// TwinCAT 3 PLC project TC3_CNCPLCBase
// Title: CNC PLC Project
// Company: Beckhoff Automation GmbH
// Author: Beckhoff Automation GmbH
// ProjectVersion: 3.1.5000.18
// Description: TwinCAT CNC Base Project
// ProgramVersion: 3.1.4026.23
// libraries:
//   Tc2_CncHli, * (Beckhoff Automation GmbH)
//   Tc2_Standard, * (Beckhoff Automation GmbH)
//   Tc2_System, * (Beckhoff Automation GmbH)
//   Tc3_CNC, * (Beckhoff Automation GmbH)
//   Tc3_EventLogger, * (Beckhoff Automation GmbH)
//   Tc3_JsonXml, * (Beckhoff Automation GmbH)
//   Tc3_Module, * (Beckhoff Automation GmbH)
// project tree:
//   CNC/ Global_CNC.TcGVL, PRG_CNCAxesHandler.TcPOU, PRG_CNCChannelHandler.TcPOU, PRG_CNCDiagnostics.TcPOU, PRG_CNCManualMode.TcPOU, PRG_CNCVariablesViewer.TcPOU, PRG_ManualFnc.TcPOU
//   / FAST.TcPOU, MAIN.TcPOU, PlcFastTask.TcTTO, PlcTask.TcTTO
//   HMI/ Global_HMI.TcGVL, ST_MachineData.TcDUT, ST_MachineMode.TcDUT, ST_MANUAL.TcDUT, ST_Position.TcDUT
//   Messages/ FB_Alarm.TcPOU, Global_Messages.TcGVL, PRG_MessagesV2.TcPOU
//   Samples/ PRG_FastMFunctions.TcPOU
// real-time tasks:
//   TASK PlcTask: cycle T#10ms, priority 20, ADS port 350
//   TASK PlcFastTask: cycle T#10ms, priority 21, ADS port 351
//   TASK CNC-Task ADS: cycle default, priority 7, ADS port 558
//   TASK CNC-Task COM: cycle T#10ms, priority 13, ADS port 556
//   TASK CNC-Task SDA: cycle T#10ms, priority 8, ADS port 555
//   TASK CNC-Task GEO: cycle T#2ms, priority 3, ADS port 554

CONFIGURATION TC3_CNCPLCBase
    RESOURCE PLC ON TwinCAT3
        TASK PlcFastTask(INTERVAL := T#10ms, PRIORITY := 21);
        TASK PlcTask(INTERVAL := T#10ms, PRIORITY := 20);
        PROGRAM FAST WITH PlcFastTask : FAST;
        PROGRAM MAIN WITH PlcTask : MAIN;
    END_RESOURCE
END_CONFIGURATION

// ---- HMI/ST_MachineData.TcDUT
TYPE ST_MachineData :
STRUCT
	// @1: Value1
	Value1: INT;
	// @1: Bool Value
	Value2: bool;
	// @1: Position
	pos : ST_Position;
	// @1: Manual @6:1
	manualFunction : ST_Manual;
END_STRUCT
END_TYPE

// ---- HMI/ST_MachineMode.TcDUT
TYPE ST_MachineMode :
STRUCT
	/// Operation Mode 
	Standby: BOOL;
	Manual: BOOL;
	MDI: BOOL;
	Automatic: BOOL;
	///REFERENCE		: BOOL;  TC3HR
	Homing: BOOL;
	/// Operation State
	Select : BOOL; 
	Ready  : BOOL;
	Start: BOOL;
	Stop: BOOL;
	Reset: BOOL;
	Error: BOOL;
	/// Special functions 
	ChannelSignals: ST_ChannelSignals;
	BlockSearch: ST_BlockSearch;
	SyntaxCheck: ST_SyntaxCheck;
	ManualMode: ST_ManualMode;
	/// Strings 
//	ProgramName: STRING(1024);
//	MDIString: STRING(1024);
	ProgramName: STRING(HLI_IMCM_MODE_STATE_PARAM_STRL);
	MDIString: STRING(HLI_IMCM_MODE_STATE_PARAM_STRL);

END_STRUCT
END_TYPE

// ---- HMI/ST_MANUAL.TcDUT
TYPE ST_MANUAL :
STRUCT
	// @1:cylinder one @2:on:1 @3:off:1 @4:pos1:1 @5:pos2:0
	cyl1 			: BYTE;	
	cyl1Status		: BYTE;
	
	// @1:conveyor @2:IMG1:1 @2:IMG2 @3:IMG15 @4:IMG16 @5:IMG7 @6:IMG13 @7:IMG14
	conv 			: BYTE;
	convStatus 		: BYTE;
	
	
END_STRUCT
END_TYPE

// ---- HMI/ST_Position.TcDUT
TYPE ST_Position :
STRUCT
	// @1:X
	x	:	LREAL;
	// @1:Y
	y	: 	LREAL;
	// @1:Z	
	Z	: 	LREAL;
END_STRUCT
END_TYPE

// ---- CNC/Global_CNC.TcGVL
VAR_GLOBAL CONSTANT
	MAX_USED_CHANNEL_IDX		: INT := 2;									(* Max index of channel that is used starting at 0, example: 1 -> totally 2 channels, maximum of 11 (12 channels) is allowed here *)
	libVersion					: ST_LibVersion := stLibVersion_Tc3_CNC;  	 
END_VAR

// ---- HMI/Global_HMI.TcGVL
VAR_GLOBAL
	/// HMI -> PLC 
	PLCChannelSignals: ST_ChannelSignals;
	/// HMI -> PLC 
	PLCSelectedChannel: INT := 0;
	/// HMI -> PLC 
	PLCFeedOverride: UINT := 100;
	/// HMI -> PLC 
	PLCSpindleOverride: UINT := 100;
	/// HMI -> PLC 
	PLCAxisEnable: BOOL;
	/// PLC -> HMI  
	PLCStatusAxisEnabled : BOOL;	
	/// HMI -> PLC 
	PLCReset: BOOL;
	PLCMachineMode: ARRAY[0..MAX_USED_CHANNEL_IDX] OF ST_MachineMode;
	/// PLC -> HMI : angewähltes File 
	PLCToHmiFile: STRING(255);
	/// Variablen für das Module "InformPlc" 
	bToggle: BOOL;
	sActualForm: STRING(255);
	nUserLevel: INT;
	sUserName: STRING(255);
	/// steigende Flanke: Applikation beenden 
	bExitApp: BOOL;	
	
	userActivity : BOOL;
	
	// @1:MachineData
	MachineData : ST_MachineData;
	
	// spindle manual mode
	nSpindleRpm:	DINT;	
	bSpindleStart: BOOL;
	bSpindleStop: BOOL;
	
	ManualFnc : ARRAY[0..3] OF FB_ManualFncFull;
	
END_VAR

// ---- Messages/Global_Messages.TcGVL
VAR_GLOBAL
	///--------------------------
	///	Messages                
	///--------------------------
	MSG_WARNING_List: ARRAY[FIRST_MESSAGE..LAST_MESSAGE] OF BOOL;
	MSG_WARNING_ListQuit: ARRAY[FIRST_MESSAGE..LAST_MESSAGE] OF BOOL;	
	MSG_ALARM_List: ARRAY[FIRST_MESSAGE..LAST_MESSAGE] OF BOOL;
	MSG_ALARM_ListQuit: ARRAY[FIRST_MESSAGE..LAST_MESSAGE] OF BOOL;			
END_VAR

VAR_GLOBAL CONSTANT
	FIRST_MESSAGE: UDINT := 1;
	LAST_MESSAGE: UDINT := 50;	
END_VAR

// ---- FAST.TcPOU
PROGRAM FAST
VAR
	nChan : INT;
	MOS_TS: INT;
	i: INT;	
	ChannelMHTFunction : ARRAY[0..MAX_USED_CHANNEL_IDX] OF HLI3_QuitChannelMHTFunction;
END_VAR

(****************************************************************************************)
(*	  							Wait for HLI initialization								*)
(****************************************************************************************)
IF NOT CNCSystem.bHLIInit THEN
	RETURN;
END_IF

IF PRG_CNCChannelHandler.stOptions.bDisableMFunctHandling THEN
	FOR i := 0 TO MAX_USED_CHANNEL_IDX DO
		ChannelMHTFunction[i](nChanIdx:=0, bM30Acknowledgement := TRUE);
	END_FOR
END_IF	

(* Programm call for MOS_TS M functions *)
// PRG_FastMFunctions();

END_PROGRAM

// ---- CNC/PRG_CNCChannelHandler.TcPOU
PROGRAM PRG_CNCChannelHandler
VAR	
	nChan					: INT;
	nOldSelectedChannel		: UDINT;
	CNCChannel				: ARRAY[0..MAX_USED_CHANNEL_IDX] OF HLI3_CNCChannel;	
	BlockSearch_Channel		: ARRAY[0..MAX_USED_CHANNEL_IDX] OF HLI3_BlockSearch;
	ErrorHandler_Channel	: ARRAY[0..MAX_USED_CHANNEL_IDX] OF FB_ChannelError;
	nChanNo: UDINT;	
	i: INT;	
	stOptions				: ST_CNC_CH_Options;
END_VAR

(****************************************************************************************)
(* POU:		PRG_ChannelHandler                     										*)
(* Type:	PRG																			*)
(* Author: 	HR / TV / MiB                                          						*)
(* Date: 	23.01.11																	*)
(* Last:	29.03.18																	*)
(* Rev.: 	1.6                                              							*)
(* ------------------------------------------------------------------------------------ *)
(* Desc:	Description																	*)
(****************************************************************************************)

(****************************************************************************************)
(*	  Map CNC function selection from HMI to selected channel (and state vice versa)  	*)
(****************************************************************************************)
IF (nOldSelectedChannel <>INT_TO_UDINT(PLCSelectedChannel)) THEN
	PLCChannelSignals.SingleBlock 		:= PLCMachineMode[PLCSelectedChannel].ChannelSignals.SingleBlock;
	PLCChannelSignals.PrgBlockIgnore	:= PLCMachineMode[PLCSelectedChannel].ChannelSignals.PrgBlockIgnore;
	PLCChannelSignals.M01Stop 			:= PLCMachineMode[PLCSelectedChannel].ChannelSignals.M01Stop;
	PLCChannelSignals.Backward 			:= PLCMachineMode[PLCSelectedChannel].ChannelSignals.Backward;
	PLCChannelSignals.FeedHold 			:= PLCMachineMode[PLCSelectedChannel].ChannelSignals.FeedHold;
	nOldSelectedChannel 				:= INT_TO_UDINT(PLCSelectedChannel);
END_IF

PLCMachineMode[PLCSelectedChannel].ChannelSignals.SingleBlock 		:= PLCChannelSignals.SingleBlock;
PLCMachineMode[PLCSelectedChannel].ChannelSignals.PrgBlockIgnore 	:= PLCChannelSignals.PrgBlockIgnore;
PLCMachineMode[PLCSelectedChannel].ChannelSignals.M01Stop 			:= PLCChannelSignals.M01Stop;
PLCMachineMode[PLCSelectedChannel].ChannelSignals.Backward 		:= PLCChannelSignals.Backward;
PLCMachineMode[PLCSelectedChannel].ChannelSignals.FeedHold 		:= PLCChannelSignals.FeedHold;


stOptions.bReferenceModeStartRequired := FALSE;

FOR i := 0 TO MAX_USED_CHANNEL_IDX DO
		
	nChan := i;	
	IF (HLI3_CheckChannelValid(nChan)) THEN		
		
		(* Error handler for channel 1 *)
		ErrorHandler_Channel[nChan](nChanIdx			:= nCHan);				
				
		(* Channel interface *)
		CNCChannel[nChan]
			(nChanIdx			:= nChan,							
			 // Operation Mode with VAR_IN_OUT Variables 
			 bModeStandby		:= PLCMachineMode[nChan].Standby,
			 bModeAutomatic		:= PLCMachineMode[nChan].Automatic,
			 bModeManual		:= PLCMachineMode[nChan].Manual,
			 bModeMDI			:= PLCMachineMode[nChan].MDI,	 
			 bModeReference		:= PLCMachineMode[nChan].Homing,
			 // Operation State with VAR_IN_OUT Variables
			 bStateSelect		:= PLCMachineMode[nChan].Select,
			 bStateReady		:= PLCMachineMode[nChan].Ready,
			 bStateStart		:= PLCMachineMode[nChan].Start,
			 bStateStop			:= PLCMachineMode[nChan].Stop,
			 bStateReset		:= PLCMachineMode[nChan].Reset,
			 // Operation Mode with VAR_IN Varaibles, the command is executed with a rising edge 
			 bCmdAutomatic 		:= FALSE,
			 bCmdManual 		:= FALSE,
    		 bCmdReference 		:= FALSE,
    		 bCmdMDI 			:= FALSE,		
			 // Operation State with VAR_IN Varaibles, the command is executed with a rising edge
			 bCmdStart 			:= FALSE,
			 bCmdStop  			:= FALSE,
	         bCmdReset 			:= FALSE,					 			 
			 // EmergencyStop 
			 bEmergencyStop 	:= FALSE,		(* If TRUE the interpolation will be aborted, Signal is no TwinSAFE function !*)
			 // Override 
			 nFeedOverride		:= PLCFeedOverride * 10,
			 nRapidFeedOverride := PLCFeedOverride * 10, 
			 // Special Functions 
			 sProgramName		:= PLCMachineMode[nChan].ProgramName,			 
			 sMDIString			:= PLCMachineMode[nChan].MDIString,
			 bBackwardMotion	:= PLCMachineMode[nChan].ChannelSignals.Backward,
			 bPrgBlockIgnore	:= PLCMachineMode[nChan].ChannelSignals.PrgBlockIgnore,
			 bFeedHold			:= PLCMachineMode[nChan].ChannelSignals.FeedHold,
			 bSingleBlock		:= PLCMachineMode[nChan].ChannelSignals.SingleBlock,
			 bDoSingleBlock		:= PLCMachineMode[nChan].ChannelSignals.DoSingleBlock,
			 bM01Stop			:= PLCMachineMode[nChan].ChannelSignals.M01Stop,
			 nSyntaxCheck		:= PLCMachineMode[nChan].SyntaxCheck.nType,
			 bM30Acknowledgement:= TRUE,
			 // Manual Mode 			 						 
			 stManualModeParameter  	 	 := stManualModeParameter[nChan],
			 stManualModeControlElements	 := stManualModeControlElements[nChan],
			 stManualModeControlElementState := stManualModeControlElementState,
			 // Options
			 stOptions			:= 	stOptions			 			 
			);
		
		(* Handle block search *)
		BlockSearch_Channel[nChan]
			(nChanIdx			:= nChan,
			 bStartRead      	:= PLCMachineMode[nChan].BlockSearch.bStartRead,   (* Edge signal *)
			 bStartWrite     	:= PLCMachineMode[nChan].BlockSearch.bStartWrite,  (* Edge signal *)
			 BlockSearch		:= PLCMachineMode[nChan].BlockSearch
			);
		
		CNCSystem.Channel[nChan].ActDistance 	:= DINT_TO_LREAL(BlockSearch_Channel[nChan].coveredDistance_AfterReset) / 10.0;
		CNCSystem.Channel[nChan].ActBlockCount 	:= BlockSearch_Channel[nChan].actualBlockCount_AfterReset;
						
	END_IF
END_FOR

END_PROGRAM

// ---- MAIN.TcPOU
PROGRAM MAIN
VAR
  
END_VAR

HLI3_Init(); 
PRG_MessagesV2();   // Messages Eventlogger V2

(* Call CNC related code only if the HLI has been initialized succesfully! *)
IF CNCSystem.bHLIInit THEN
	PRG_CNCAxesHandler();    	
	PRG_CNCManualMode();
	PRG_CNCChannelHandler();	
	PRG_CNCVariablesViewer();
	PRG_ManualFnc();
	PRG_CNCDiagnostics();		
END_IF
(* Reset the reset flag from HMI *)
PLCReset := FALSE;

END_PROGRAM

// ---- Messages/PRG_MessagesV2.TcPOU
PROGRAM PRG_MessagesV2
VAR
	arrAlarmSimple: ARRAY[1..10] OF FB_Alarm;	
	bTestAlarm1: BOOL;
	bTestAlarm2: BOOL;
	bTestAlarm3: BOOL;
	sTestString : STRING := 'this is a test line';
END_VAR

;

(* add Alarms.tmc to "Systen\Type System" before uncommenting this *)

(*
arrAlarmSimple[1](Event := TC_EVENTS.Alarms.Alarm1);
arrAlarmSimple[1].Raise := bTestAlarm1;
arrAlarmSimple[1].AddInfo := sTestString;


arrAlarmSimple[2](Event := TC_EVENTS.Alarms.Alarm2);
arrAlarmSimple[2].Raise := bTestAlarm2;

arrAlarmSimple[3](Event := TC_EVENTS.Alarms.Alarm3);
arrAlarmSimple[3].Raise := bTestAlarm3;
*)

END_PROGRAM

// ---- Messages/FB_Alarm.TcPOU
FUNCTION_BLOCK FB_Alarm
VAR_INPUT
	Event : TcEventEntry;  // AlarmEntry from TMS Editor. Example: TC_EVENTS.Alarms.Alarm1
	Raise : BOOL;		   // true -> Alarm is active, false -> Alarm not active
	AddInfo: STRING;	   // if <> empty -> additional Info that is transfered together with alarm
END_VAR
VAR_OUTPUT
END_VAR
VAR
	_alarm : FB_TcAlarm;
	_initDone : BOOL;
	_rTrigRaise : R_TRIG;
	_fTrigRaise : F_TRIG;
	_fbSourceInfo : FB_TcSourceInfo;
	_fbJson      : FB_JsonSaxWriter;
	_sJsonDoc    : STRING(255);	
END_VAR

(* ========================================================= *)
(*    FUN: FB_Alarm                   					     *)
(* --------------------------------------------------------- *)
(*   Desc: Simple usage of Eventlogger2 Alarms               *)
(* Author: MiB                                               *)
(*   Date: 09.03.2021                                        *)
(*   Rev.: 1.0                                               *)
(* ========================================================= *)


// init
IF NOT _initDone AND Event.nEventId <> 0 THEN
	_fbSourceInfo.sName := 'PLC';
	_alarm.CreateEx(Event, FALSE, _fbSourceInfo );
	_initDone := TRUE;
END_IF

// raise alarm
_rTrigRaise(clk := Raise);
IF _rTrigRaise.Q AND NOT _alarm.bRaised  THEN
	IF LEN(AddInfo) > 0 THEN 
		_fbJson.ResetDocument();
		_fbJson.StartObject();
		_fbJson.AddKey('AddInfo');
		_fbJson.AddString(AddInfo);		
		_fbJson.EndObject();
		_sJsonDoc := _fbJson.GetDocument();
	    _alarm.SetJsonAttribute(_sJsonDoc);		
	ELSE
		_alarm.SetJsonAttribute('');
	END_IF
	_alarm.Raise(0);
END_IF

// clear alarm
_fTrigRaise(clk := Raise);
IF _fTrigRaise.Q AND _alarm.bRaised THEN
	_alarm.Clear(0, FALSE);
END_IF

END_FUNCTION_BLOCK

// ---- CNC/PRG_CNCAxesHandler.TcPOU
PROGRAM PRG_CNCAxesHandler
VAR
	nHliAxisIdx					: INT;				
	fbCNC_Axis					: ARRAY[0..HLI_SYS_AX_MAXIDX] OF FB_CNCAxis;	
	
	nFirstSpindle				: INT := -1;
	fbHandleSpindleTechno		: HLI3_HandleSpindleTechnoGearChange;
	M3,M4,M5,M19				: BOOL;
	MDummy						: BOOL;
	M40, M41, M42, M43, M44, M45: BOOL;
	
	fbHandleSpindleTechno2		: HLI3_HandleSpindleTechno;
	M3_1,M4_1,M5_1,M19_1				: BOOL;
	
	
	fbAxesError 				: FB_AxesError;
		
	// FB_CNCAxis Sample
	// fbAxis_X 					:  FB_CNCAxis; 
	// stParameter					:  ST_CNC_AX_Parameter;
	// stOptions					:  ST_CNC_AX_Options;
	// stPLCopen					:  ST_CNC_AX_PLCopen;
			
	(*
	fbHandleSpindleTechnoPlcSp	: HLI3_HandleSpindleTechno;
	SM3,SM4,SM5,SM19			: bool; 
	*)
	bCalibrationCam: BOOL;
	fbMoveSpindle: HLI3_MoveSpindle;
	

	
	probingSignal: BOOL;
	
	SpindleControl: ST_SpindleControl;
	fbMoveSpindle2: HLI3_MoveSpindleControl;
	rTrigReset : R_TRIG;
END_VAR

(****************************************************************************************)
(* POU:		PRG_AxesHandler                     										*)
(* Type:	PRG																			*)
(* Author: 	TV,MiB                                             							*)
(* Date: 	20.02.2019																	*)
(* Rev.: 	1.6                                               							*)
(* ------------------------------------------------------------------------------------ *)
(* Desc:	Description																	*)
(****************************************************************************************)

fbAxesError(bReset := PLCReset);

(****************************************************************************************)
(*							Release of all reachable axes								*)
(****************************************************************************************)
PLCStatusAxisEnabled := TRUE;   
FOR nHliAxisIdx := 0 TO UDINT_TO_INT(gNrAx-1) DO			
	fbCNC_Axis[nHliAxisIdx](
		nLogAxisNo :=  UINT_TO_INT(gpAx[nHliAxisIdx]^.head.log_ax_nr_r),
		bEnable		:= PLCAxisEnable AND (nHliAxisIdx <> 1));
		IF (NOT fbCNC_Axis[nHliAxisIdx].stStatus.bIsEnabled) THEN    // if one axis status is "not enabled" -> reset PLCStatusAxisEnabled
			PLCStatusAxisEnabled := FALSE;
		END_IF
		IF HLI3_CheckAxisValid(nHliAxisIdx) THEN
			IF nFirstSpindle = -1 AND gpAx[nHliAxisIdx]^.ipo_state.spindle_axis_r THEN  (* store HLIIndex of first spindle *)
				nFirstSpindle := nHliAxisIdx;
			END_IF
		END_IF
END_FOR
fbCNC_Axis[0].stOptions.bDisableAutoFollowUp := TRUE;

fbCNC_Axis[0].stOptions.bProbingSignal := probingSignal;



	// FB_CNCAxis Sample 

	// CNC Axis Options
	
	// stOptions.strPathCompTable;
	// stOptions.bActivateCompTable;
	// stOptions.bProbingSignal;
	// stOptions.bReducedSpeed;
	// stOptions.bReducedSpeedZone1;
	// stOptions.bReducedSpeedZone2;
	// stOptions.bResetCalibration;
	
	// CNC Parameters
			
	// stParameter.bWriteParameter;
	// stParameter.nNumParameters  	:= 2;
	// stParameter.strTempPath		:= 'C:\';
	
	// stParameter.ParamList[0].strName 	:= 'kenngr.swe_pos';
	// stParameter.ParamList[0].strValue 	:= '30000000';

	// stParameter.ParamList[1].strName 	:= 'kenngr.swe_neg';
	// stParameter.ParamList[1].strValue 	:= '0';

	// PLCOpen
	// stPLCopen.nOverride;
	// stPLCopen.bExecuteHoming;
	// stPLCopen.bCamSignal;
	// stPLCopen.bExecuteMoveAbsolute;
	// stPLCopen.bExecuteReset;
	// stPLCopen.fPosition;
	// stPLCopen.fVelocity;
	// stPLCopen.fAcceleration;
	// stPLCopen.fJerk;
	
	(*
	fbAxis_X(
		nLogAxisNo:=1, 
		bEnable:= PLCAxisEnable, 
		bCalibrationCam:= bCalibrationCam, 
		bSetRefOffset:= , 
		fRefOffset:= , 
		bFeedhold:= ,
		stOptions:= stOptions, 
		stParameter:= stParameter, 
		stPLCopen:= stPLCopen, 
		stStatus=> );
*)		
 




	fbHandleSpindleTechno2(
		nHliAxisIdx:=15 , 		
		bIsChannelSpecific:= FALSE, 
		bHandleGearChange := FALSE,		
		nRevolution=> , 
		nPosition=> , 
		bError=> , 
		nErrorId=> , 
		M03:= M3_1, 
		M04:= M4_1, 
		M05:= M5_1, 
		M19:= M19_1
		); 

	(* acknowledge all spindle M funnctions immediately *)
	M3_1 := FALSE;  
	M4_1 := FALSE;
	M5_1 := FALSE;
	M19_1 := FALSE;
	


(* if there exits spindles use the first one for spindleoverride *)
IF nFirstSpindle <> -1 THEN
	HLI3_SetAxisOverride(nHliAxisIdx:= nFirstSpindle , nOverride:= PLCSpindleOverride *10);

	fbHandleSpindleTechno(
		nHliAxisIdx:=nFirstSpindle , 		
		bIsChannelSpecific:= FALSE, 
		bHandleGearChange := FALSE,		
		nRevolution=> , 
		nPosition=> , 
		bError=> , 
		nErrorId=> , 
		M03:= M3, 
		M04:= M4, 
		M05:= M5, 
		M19:= M19,
		M40 := M40,
		M41 := M41,
		M42 := M42,
		M43 := M43,
		M44 := M44,
		M45 := M45,
		); 
	(* acknowledge all spindle M funnctions immediately *)
	M3 := FALSE;  
	M4 := FALSE;
	M5 := FALSE;
	M19 := FALSE;
	
	
	
	(* Example for starting and stopping a spindle in manual mode in first channel *)
	IF (CNCSystem.Channel[0].ActMode = HLI_IMCM_MANUAL_MODE) THEN 	
		fbMoveSpindle(
			nHliAxisIdx:=nFirstSpindle , 
			nSpeed:= nSpindleRpm ,   (* defined in Global_HMI *)
			bStart:=bSpindleStart, 	 (* defined in Global_HMI *)
			bStop:= bSpindleStop , 	 (* defined in Global_HMI *)
			bBusy=> , 
			bError=> , 
			nErrID=> , 
			sErrText=> );
	END_IF
	IF (bSpindleStart AND NOT fbMoveSpindle.bBusy) THEN 
		bSpindleStart := FALSE;
	END_IF
	IF (bSpindleStop AND NOT fbMoveSpindle.bBusy) THEN 
		bSpindleStop := FALSE;
	END_IF	
	
	
END_IF



(* spindle controlling form HMI *)
FOR nHliAxisIdx := 0 TO UDINT_TO_INT(gNrAx-1) DO			
	IF gpAx[nHliAxisIdx]^.ipo_state.spindle_axis_r  THEN
		HLI3_SetAxisOverride(nHliAxisIdx:= nHliAxisIdx , nOverride:= PLCSpindleOverride *10);
	END_IF	
END_FOR

rTrigReset(clk := PLCReset);
IF rTrigReset.Q THEN
	SpindleControl.busy := FALSE;
END_IF

fbMoveSpindle2(
    stControl   := SpindleControl,
	bReset		:= PLCReset,
    bBusy       => ,
    bError      => ,
    nErrID      => ,	
    sErrText    => );



(* Howto use plc controlled spindle : *)
(*
fbHandleSpindleTechnoPlcSp(
	nHliAxisIdx:= 0 , 
	nHliChannelIdx:= 0 , 
	bIsChannelSpecific:= TRUE, 
	nLogAxisNoChannelSpecific:= 95 , 
	bHandleGearChange:= FALSE , 
	bChannelReset:= FALSE, 
	nRevolution=> , 
	nPosition=> , 
	bError=> , 
	nErrorId=> , 
	M03:= SM3, 
	M04:= SM4, 
	M05:= SM5, 
	M19:= SM19);
*)

END_PROGRAM

// ---- CNC/PRG_CNCManualMode.TcPOU
PROGRAM PRG_CNCManualMode
VAR
	fbUintUdInt: ARRAY [0..MAX_USED_CHANNEL_IDX] OF FB_Uint_Udint;
	nHandwheel : UINT;		(* increments for handwheel (e.g. EL5101   *)
	nHandWheelBig: UDINT;
	i: INT;
END_VAR


FOR i := 0 TO MAX_USED_CHANNEL_IDX DO
	
	IF (HLI3_CheckChannelValid(i)) THEN

		stManualModeParameter[i].stChannelParameter.nChanIdx						:= i;       (* Channel 1 *)
		stManualModeParameter[i].stChannelParameter.nInc							:= PLCMachineMode[i].ManualMode.nInc * 10;
		stManualModeParameter[i].stChannelParameter.bG200ConfigurationViaPLC		:= TRUE;		
		
		stManualModeParameter[i].stChannelParameter.eManualType						:= UINT_TO_INT(PLCMachineMode[i].ManualMode.nManualTyp);			
		IF (stManualModeParameter[i].stChannelParameter.eManualType = E_CNC_ManualType.Handwheel AND i <> PLCSelectedChannel) THEN	(* if in Handwheel mode and the channel is NOT selected -> leave handwheel mode and change to TippMode*)
			stManualModeParameter[i].stChannelParameter.eManualType						:= E_CNC_ManualType.TippMode;
		END_IF		
		
		stManualModeParameter[i].stChannelParameter.stManualOption.bTrafoActive := PLCMachineMode[i].ManualMode.stManualOption.bTrafoActive;
        stManualModeParameter[i].stChannelParameter.stManualOption.bEcsActive := PLCMachineMode[i].ManualMode.stManualOption.bEcsActive;
        stManualModeParameter[i].stChannelParameter.stManualOption.eZeroOffset := PLCMachineMode[i].ManualMode.stManualOption.eZeroOffset;
							
		
		stManualModeParameter[i].stChannelParameter.nHandwheelResolution			:= UDINT_TO_DINT(PLCMachineMode[i].ManualMode.nHwResolution);    (* 0.1 µm /rev (from HMI) *)						
		stManualModeParameter[i].stAxisParameter.stControlUnit[0].nLogAxisNr		:= PLCMachineMode[i].ManualMode.nLogAxisNumber;   (* Log. Achs Nummer *)
		IF stManualModeParameter[i].stAxisParameter.stControlUnit[0].nLogAxisNr = 0 THEN
			stManualModeParameter[i].stAxisParameter.stControlUnit[0].nLogAxisNr := gpCh[i]^.bahn_state.coord_r[0].log_achs_nr_r;
			PLCMachineMode[i].ManualMode.nLogAxisNumber := gpCh[i]^.bahn_state.coord_r[0].log_achs_nr_r;
		END_IF
		stManualModeParameter[i].stAxisParameter.stControlUnit[0].nSpeed			:= LREAL_TO_UDINT(PLCMachineMode[i].ManualMode.nSpeed * 16.666);
		stManualModeControlElements[i].stControlKeys[0].bKeyNeg						:= PLCMachineMode[i].ManualMode.bKeyNeg;
		stManualModeControlElements[i].stControlKeys[0].bKeyPos						:= PLCMachineMode[i].ManualMode.bKeyPos;
		stManualModeControlElements[i].stControlKeys[0].bKeyRapid					:= PLCMachineMode[i].ManualMode.bKeyRapid;
		
		(* the cnc needs an UDINT for handwheel increments, fbUintUdint extends an UInt to an UDINT *)
		(* the resoltion of the handwheel is parameterized in CNC-Task GEO/Manual MDS: (e.g. 400 handwheel inc / handwheel revolution
		
				hr_data[0].hr_aufl_z              400         ( P-MANU-00005 : Handwheel resolution numerator
				hr_data[0].hr_aufl_n                1     	  ( P-MANU-00006 : Handwheel resolution denominator
		*) 
		fbUintUdInt[i](nInSmall := nHandwheel, nBig := nHandWheelBig);
		stManualModeControlElements[i].nHandwheelInc[0] :=  UDINT_TO_DINT(nHandWheelBig);
  END_IF
END_FOR

END_PROGRAM

// ---- CNC/PRG_CNCVariablesViewer.TcPOU
PROGRAM PRG_CNCVariablesViewer
VAR			
	fbReadCNCVariables : FB_ReadCNCVariables;		
END_VAR

fbReadCNCVariables(
	bEnable:= TRUE, 
	nChanIdx:= PLCSelectedChannel, 
	eVariablesType:= eVariablesType, 
	tIntervall:= T#1S, 	 
	stCNCVariablesViewer_Data:= stCNCVariablesViewer_Data);

END_PROGRAM

// ---- CNC/PRG_ManualFnc.TcPOU
PROGRAM PRG_ManualFnc
VAR
END_VAR



	ManualFnc[0].headerText := 'HeaderText 1';
	ManualFnc[0].addText := 'addText';
	ManualFnc[0].infoText1 := 'infoText1';
	ManualFnc[0].infoText2 := 'infoText2';
	ManualFnc[0].infoText3 := 'infoText3';
	ManualFnc[0].infoText4 := 'infoText4';
	ManualFnc[0].error := FALSE;
	
	ManualFnc[0].left.key.text := 'left.key.text';
	ManualFnc[0].left.status.text := 'left.status.text';
	ManualFnc[0].left.key.disable := TRUE;
	ManualFnc[0].left.status.colorChange := TRUE;
	
	ManualFnc[0].right.key.text := 'right.key.text';
	ManualFnc[0].right.status.text := 'right.status.text';
	ManualFnc[0].right.key.colorChange := TRUE;

	
	

	ManualFnc[1].headerText := 'HeaderText 2';
	ManualFnc[1].addText := '';
	ManualFnc[1].infoText1 := 'infoText1';
	ManualFnc[1].infoText2 := 'infoText2';
	ManualFnc[1].infoText3 := 'infoText3';
	ManualFnc[1].infoText4 := 'infoText4';
	ManualFnc[1].error := FALSE;
	ManualFnc[1].select := FALSE;
		
	ManualFnc[1].left.key.text := 'left.key.text';
	ManualFnc[1].left.status.text := 'left.status.text';
	ManualFnc[1].left.key.disable := FALSE;
	ManualFnc[1].left.status.colorChange := FALSE;
	
	ManualFnc[1].right.key.text := 'right.key.text';
	ManualFnc[1].right.status.text := 'right.status.text';
	ManualFnc[1].right.key.colorChange := FALSE;
	



	
	ManualFnc[2].headerText := 'HeaderText 3';
	ManualFnc[2].addText := 'addText';
	ManualFnc[2].infoText1 := 'infoText1';
	ManualFnc[2].infoText2 := 'infoText2';
	ManualFnc[2].infoText3 := 'infoText3';
	ManualFnc[2].infoText4 := 'infoText4';
	ManualFnc[2].error := TRUE;
	
	ManualFnc[2].left.key.text := 'left.key.text';
	ManualFnc[2].left.status.text := 'left.status.text';
	ManualFnc[2].left.key.disable := TRUE;
	ManualFnc[2].left.status.colorChange := TRUE;
	
	ManualFnc[2].right.key.text := 'right.key.text';
	ManualFnc[2].right.status.text := 'right.status.text';
	ManualFnc[2].right.key.colorChange := TRUE;	
	


	
	
	ManualFnc[3].headerText := 'HeaderText 4';
	ManualFnc[3].addText := '';
	ManualFnc[3].infoText1 := 'infoText1';
	ManualFnc[3].infoText2 := 'infoText2';
	ManualFnc[3].infoText3 := 'infoText3';
	ManualFnc[3].infoText4 := 'infoText4';
	ManualFnc[3].error := FALSE;
	ManualFnc[3].select := FALSE;	
	
	ManualFnc[3].left.key.text := 'left.key.text';
	ManualFnc[3].left.status.text := 'left.status.text';
	ManualFnc[3].left.key.disable := FALSE;
	ManualFnc[3].left.status.colorChange := FALSE;
	
	ManualFnc[3].right.key.text := 'right.key.text';
	ManualFnc[3].right.status.text := 'right.status.text';
	ManualFnc[3].right.key.colorChange := FALSE;

END_PROGRAM

// ---- CNC/PRG_CNCDiagnostics.TcPOU
PROGRAM PRG_CNCDiagnostics
VAR
	fbCNCDiagnosisUpload : FB_CNCDiagnosisUpload;
	bUploadDiagData: BOOL;
END_VAR

fbCNCDiagnosisUpload(
	bExecute:= bUploadDiagData, 
	strFileName:= 'C:\temp\diag_data.txt', 
	nHistory:= 0, 
	strTopic:= 'ALL', 
	bBusy=> , 
	bError=> , 
	nErrorID=> );

END_PROGRAM

// ---- Samples/PRG_FastMFunctions.TcPOU
PROGRAM PRG_FastMFunctions
VAR
	anMFunctionNo						: ARRAY[0..MAX_FAST_M_FUNC_ITEM_IDX] OF UINT;	
	fbFastMFunctionProvider				: HLI3_FastMFunctionProvider;
	fbFastMFunctionHandler				: HLI3_FastMFunctionHandler;	
	abyOutput					AT %Q*	: ARRAY[0..MAX_FAST_M_FUNC_OUTPUT_IDX] OF BYTE;  	
END_VAR

(****************************************************************************************)
(* POU:		PRG_FastMFunctions                    										*)
(* Type:	PRG																			*)
(* Author: 	RCH		                                             						*)
(* Date: 	14/10/29																	*)
(* Rev.: 	1.0                                               							*)
(* ------------------------------------------------------------------------------------ *)
(* Desc.:	PLC program to demonstrate usage of MOS_TS M functions using the FB´s		*)
(*			HLI3_FastMFunctionProvider and HLI3_FastMFunctionHandler.					*)
(*			In order to achieve a determenistic output behavior this program has to be 	*)
(*			called by a task running synchronously to the CNC GEO task. Therefore that	*)
(*			task´s priority  has to be adjusted in a way that it gets called by the 	*)
(* 			realtime system	right after the CNC GEO task.								*)
(*																						*)
(*			THIS IMPLEMENTATION REQUIRES A 1MS CNC GEO AND 1MS FAST PLC TASK CYCLE!!!	*)
(* ------------------------------------------------------------------------------------ *)
(* Rev.:	<Enter revision number here>												*)
(* Date:	<Enter revision data here>				                                   	*)
(* Author:	<Enter author´s shortcut here>											 	*)
(* Desc.:	<Enter description here>													*)
(****************************************************************************************)


(****************************************************************************************)
(*	  						Configure M function no´s to provide						*)
(****************************************************************************************)
(* Add up to MAX_FAST_M_FUNC_ITEM_IDX m function numbers that should be handled by 		*)
(* fbFastMFunctionProvider.																*)
anMFunctionNo[0]	:= 25;
anMFunctionNo[1]	:= 26;

fbFastMFunctionProvider
	(nHliChanIdx	:= 0, 
	 anMFunctionNo	:= anMFunctionNo
	);
	
(****************************************************************************************)
(*	  						 	Handle Laser ON/OFF (M25/M26)							*)
(****************************************************************************************)
(* M function numbers for switching ON and OFF have to be contained in the 				*)
(* 'anMFunctionNo' array of the HLI3_FastMFunctionProvider instance which provides the	*)
(* 'stData' structure to this FB.														*)
(* The delay times nDelayOn and nDelayOff can be used to adopt to external hardware		*)
(* delays!																				*)
fbFastMFunctionHandler
	(bForceOff		:= FALSE, 
	 bReset			:= FALSE, 
	 nFunctionNoOn	:= 25, 
	 nDelayOn		:= 0,			
	 nFunctionNoOff	:= 26, 
	 nDelayOff		:= 0,
	 stData			:= fbFastMFunctionProvider.stData,
	 abyOutput		=> abyOutput
	);

END_PROGRAM
